FUNCTION_BLOCK EL_LinearAxis (* The logic of an equipment block: one holder at a time, outputs switched off before new ones go on, all off on release or abort, inputs reported when they change. Technical: LinearAxis: output values from its holder -> outputs (break before make); one holder at a time; all off on release or when the module aborts; inputs -> state channel when they change *)
  (* Standard: 61499-2 *)
  (* Version 0.1, 2026-09-28, Project contributors, AAU Smart Production Lab *)
  PACKAGE stoppering;
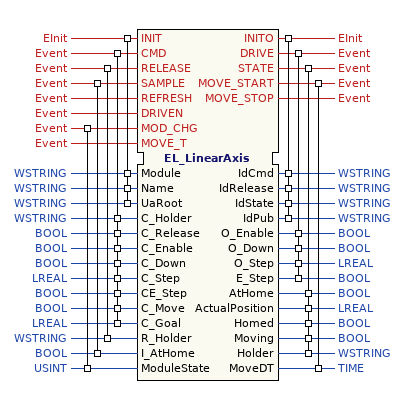
  EVENT_INPUT
    INIT : EInit WITH Module, Name, UaRoot; (* Initialise, once at start-up (the INIT chain); takes the values given with it *)
    CMD WITH C_Holder, C_Release, C_Enable, C_Down, C_Step, CE_Step, C_Move, C_Goal; (* A command arrived from a holder *)
    RELEASE WITH R_Holder; (* A release arrived on the module's release channel (R_Holder) *)
    SAMPLE WITH I_AtHome; (* The inputs were read *)
    REFRESH; (* Cycle: write the outputs again *)
    DRIVEN; (* The outputs were written *)
    MOD_CHG WITH ModuleState; (* The module's state changed (its Aborting switches all off) *)
    MOVE_T; (* The move's time is up: the axis is at the goal *)
  END_EVENT
  EVENT_OUTPUT
    INITO : EInit WITH IdCmd, IdRelease, IdState, IdPub; (* Initialised: the next block of the INIT chain goes on *)
    DRIVE WITH O_Enable, O_Down, O_Step, E_Step; (* Write the outputs *)
    STATE WITH AtHome, ActualPosition, Homed, Moving, Holder; (* Publish the state (the inputs and the holder) *)
    MOVE_START WITH MoveDT; (* Start the move's timer (MoveDT) *)
    MOVE_STOP; (* Stop the move's timer *)
  END_EVENT
  VAR_INPUT
    Module : WSTRING; (* The module's name; its local channels are named after it (loc[<Module>/...]) *)
    Name : WSTRING; (* The equipment item's name: its local channels and OPC UA folder *)
    UaRoot : WSTRING; (* The module's OPC UA folder, e.g. /Objects/Filling *)
    C_Holder : WSTRING; (* Who sends the command *)
    C_Release : BOOL; (* Give up the equipment after this command *)
    C_Enable : BOOL; (* Commanded value of Enable *)
    C_Down : BOOL; (* Commanded value of Down *)
    C_Step : LREAL; (* Commanded value of Step *)
    CE_Step : BOOL; (* Commanded: Step enabled *)
    C_Move : BOOL; (* Move to a position *)
    C_Goal : LREAL; (* The position to move to *)
    R_Holder : WSTRING; (* Who gives up the equipment *)
    I_AtHome : BOOL; (* AtHome as read or received *)
    ModuleState : USINT; (* PackML state: 1 Clearing, 2 Stopped, 3 Starting, 4 Idle, 6 Execute, 7 Stopping, 8 Aborting, 9 Aborted, 15 Resetting *)
  END_VAR
  VAR_OUTPUT
    IdCmd : WSTRING; (* Local channel of the commands *)
    IdRelease : WSTRING; (* Local channel of the releases (the module's, one for all equipment) *)
    IdState : WSTRING; (* Local channel of the state *)
    IdPub : WSTRING; (* OPC UA ID of the published inputs *)
    O_Enable : BOOL; (* The value to write to Enable *)
    O_Down : BOOL; (* The value to write to Down *)
    O_Step : LREAL; (* The value to write to Step *)
    E_Step : BOOL; (* Step enabled (FALSE writes 0) *)
    AtHome : BOOL; (* LinearAxis: AtHome, an input *)
    ActualPosition : LREAL; (* LinearAxis: ActualPosition (mm), worked out by the equipment *)
    Homed : BOOL; (* LinearAxis: Homed, worked out by the equipment *)
    Moving : BOOL; (* LinearAxis: Moving, worked out by the equipment *)
    Holder : WSTRING; (* Who holds the equipment (empty: free) *)
    MoveDT : TIME; (* How long the move takes *)
  END_VAR
  VAR
    Publish : BOOL;
    Beat : USINT;
    LastHolder : WSTRING;
    Pending : BOOL;
    OffPending : BOOL;
    L_AtHome : BOOL;
    L_Homed : BOOL;
    L_Moving : BOOL;
    N_Enable : BOOL;
    N_Down : BOOL;
    N_Step : LREAL;
    NE_Step : BOOL;
    N_Move : BOOL;
    N_Goal : LREAL;
    MoveGoal : LREAL;
    MoveFrom : LREAL;
    MoveDir : LREAL;
    MoveSince : TIME;
    MoveStart : BOOL;
    Uncounted : BOOL;
  END_VAR
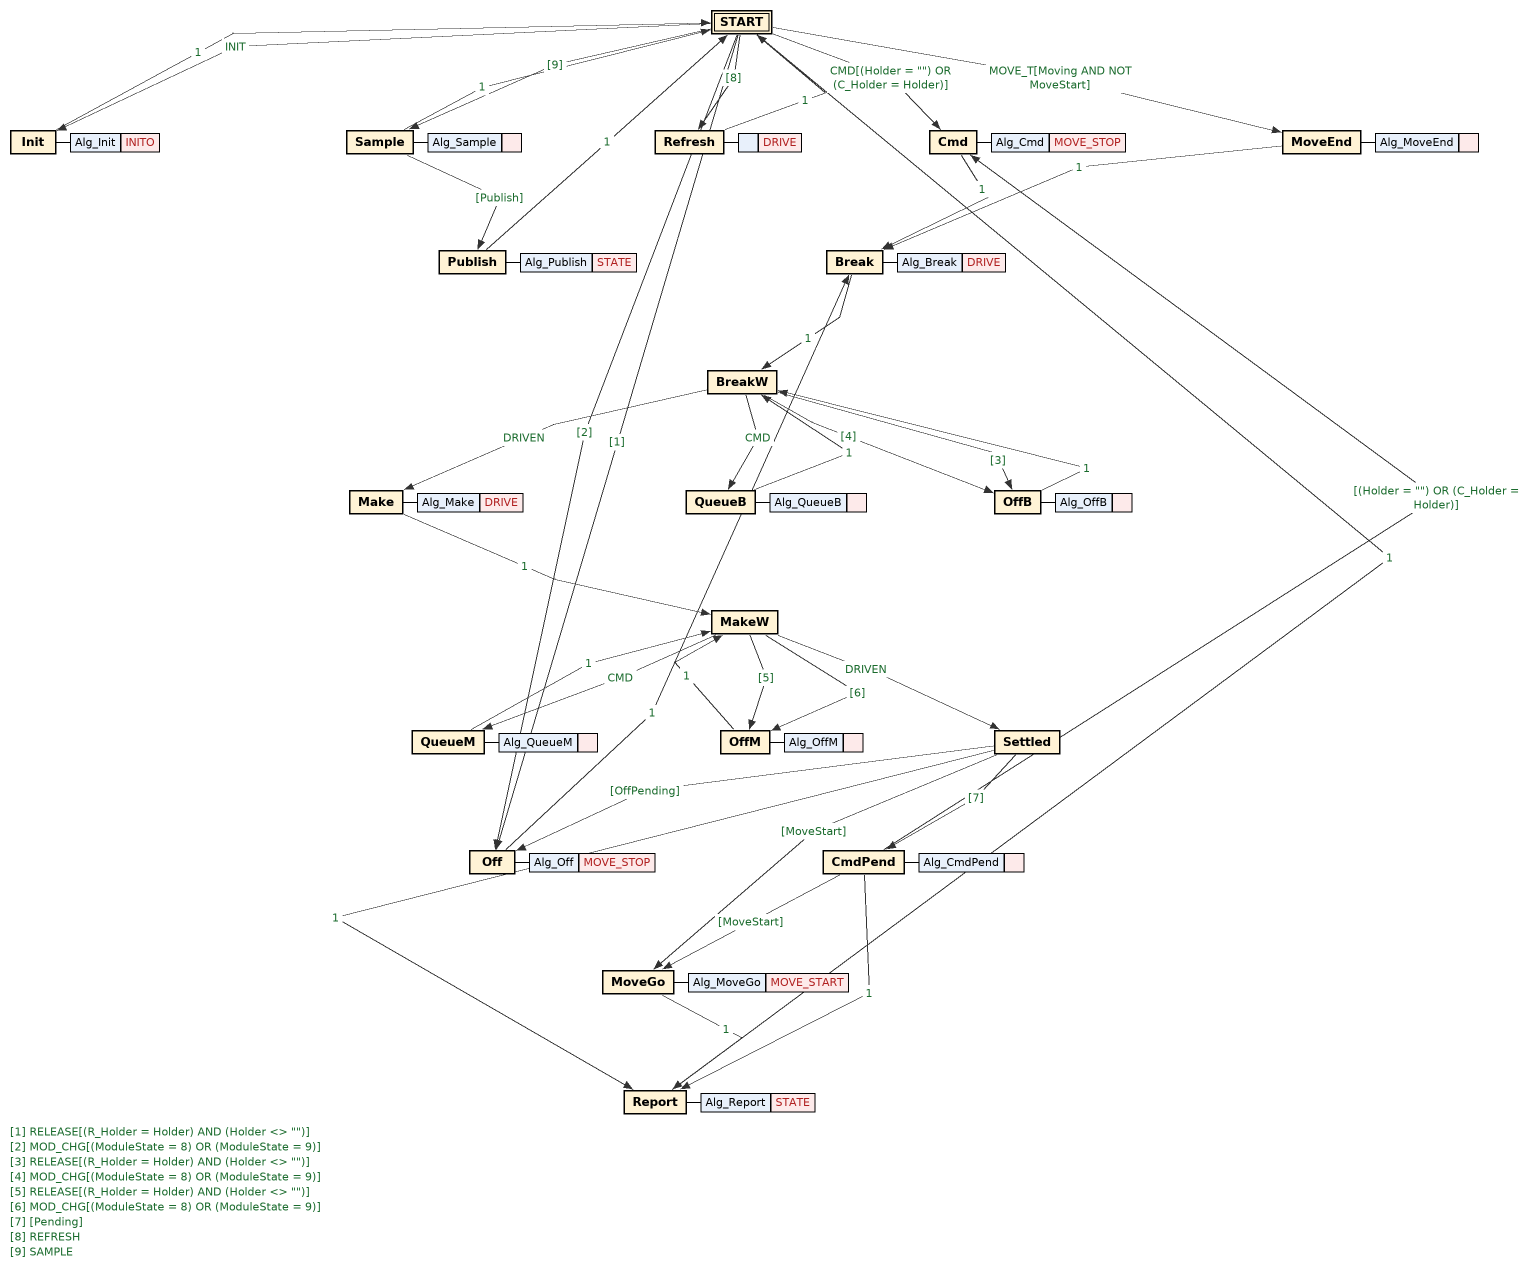
  EC_STATES
    START;
    Init : Alg_Init -> INITO;
    Sample : Alg_Sample;
    Publish : Alg_Publish -> STATE;
    Refresh : -> DRIVE;
    Cmd : Alg_Cmd -> MOVE_STOP;
    Off : Alg_Off -> MOVE_STOP;
    Break : Alg_Break -> DRIVE;
    Make : Alg_Make -> DRIVE;
    BreakW;
    MakeW;
    QueueB : Alg_QueueB;
    OffB : Alg_OffB;
    QueueM : Alg_QueueM;
    OffM : Alg_OffM;
    CmdPend : Alg_CmdPend;
    Settled;
    MoveGo : Alg_MoveGo -> MOVE_START;
    MoveEnd : Alg_MoveEnd;
    Report : Alg_Report -> STATE;
  END_STATES
  EC_TRANSITIONS
    START TO Init := INIT;
    START TO Sample := SAMPLE;
    START TO Refresh := REFRESH;
    START TO Cmd := CMD[(Holder = "") OR (C_Holder = Holder)];
    START TO Off := RELEASE[(R_Holder = Holder) AND (Holder <> "")];
    START TO Off := MOD_CHG[(ModuleState = 8) OR (ModuleState = 9)];
    START TO MoveEnd := MOVE_T[Moving AND NOT MoveStart];
    MoveEnd TO Break := 1;
    Init TO START := 1;
    Sample TO Publish := [Publish];
    Sample TO START := 1;
    Publish TO START := 1;
    Refresh TO START := 1;
    Cmd TO Break := 1;
    Off TO Break := 1;
    Break TO BreakW := 1;
    BreakW TO Make := DRIVEN;
    Make TO MakeW := 1;
    MakeW TO Settled := DRIVEN;
    BreakW TO QueueB := CMD;
    BreakW TO OffB := RELEASE[(R_Holder = Holder) AND (Holder <> "")];
    BreakW TO OffB := MOD_CHG[(ModuleState = 8) OR (ModuleState = 9)];
    QueueB TO BreakW := 1;
    OffB TO BreakW := 1;
    MakeW TO QueueM := CMD;
    MakeW TO OffM := RELEASE[(R_Holder = Holder) AND (Holder <> "")];
    MakeW TO OffM := MOD_CHG[(ModuleState = 8) OR (ModuleState = 9)];
    QueueM TO MakeW := 1;
    OffM TO MakeW := 1;
    Settled TO Off := [OffPending];
    Settled TO CmdPend := [Pending];
    CmdPend TO Cmd := [(Holder = "") OR (C_Holder = Holder)];
    CmdPend TO MoveGo := [MoveStart];
    Settled TO MoveGo := [MoveStart];
    MoveGo TO Report := 1;
    CmdPend TO Report := 1;
    Settled TO Report := 1;
    Report TO START := 1;
  END_TRANSITIONS
  ALGORITHM Alg_Init IN ST:
IdCmd := CONCAT(CONCAT(CONCAT(CONCAT("loc[", Module), "/"), Name), "/cmd]");
IdRelease := CONCAT(CONCAT("loc[", Module), "/release]");
IdState := CONCAT(CONCAT(CONCAT(CONCAT("loc[", Module), "/"), Name), "/state]");
IdPub := CONCAT(CONCAT(CONCAT(CONCAT(CONCAT(CONCAT(CONCAT(CONCAT(CONCAT(CONCAT(CONCAT(CONCAT(CONCAT(CONCAT(CONCAT(CONCAT(CONCAT("opc_ua[WRITE;", UaRoot), "/Equipment/"), Name), "/AtHome;"), UaRoot), "/Equipment/"), Name), "/ActualPosition;"), UaRoot), "/Equipment/"), Name), "/Homed;"), UaRoot), "/Equipment/"), Name), "/Moving"), "]");
  END_ALGORITHM
  ALGORITHM Alg_Sample IN ST:
AtHome := I_AtHome;
IF Moving AND NOT MoveStart THEN
  ActualPosition := MoveFrom + MoveDir * 20.0 * TIME_IN_MS_TO_LREAL(NOW_MONOTONIC() - MoveSince) / 1000.0;
  IF MoveDir * (ActualPosition - MoveGoal) > 0.0 THEN
    ActualPosition := MoveGoal;
  END_IF;
ELSIF AtHome THEN
  ActualPosition := 0.0;
  Homed := TRUE;
ELSIF Uncounted THEN
  Homed := FALSE;
END_IF;
Publish := (AtHome <> L_AtHome) OR (Homed <> L_Homed) OR (Moving <> L_Moving) OR (Holder <> LastHolder) OR (Beat >= 20) OR (Moving AND (Beat >= 4));
Beat := Beat + 1;
  END_ALGORITHM
  ALGORITHM Alg_Publish IN ST:
L_AtHome := AtHome;
L_Homed := Homed;
L_Moving := Moving;
LastHolder := Holder;
Beat := 0;
  END_ALGORITHM
  ALGORITHM Alg_Cmd IN ST:
Holder := C_Holder;
N_Enable := C_Enable;
N_Down := C_Down;
N_Step := C_Step;
NE_Step := CE_Step;
N_Move := C_Move;
N_Goal := C_Goal;
IF Moving AND NOT MoveStart THEN
  ActualPosition := MoveFrom + MoveDir * 20.0 * TIME_IN_MS_TO_LREAL(NOW_MONOTONIC() - MoveSince) / 1000.0;
  IF MoveDir * (ActualPosition - MoveGoal) > 0.0 THEN
    ActualPosition := MoveGoal;
  END_IF;
END_IF;
Moving := FALSE;
MoveStart := FALSE;
IF N_Move THEN
  IF Homed AND (ABS(N_Goal - ActualPosition) >= 0.0005) THEN
    MoveGoal := N_Goal;
    MoveFrom := ActualPosition;
    MoveDT := MUL_TIME(T#1s, ABS(N_Goal - ActualPosition) / 20.0);
    IF N_Goal > ActualPosition THEN
      MoveDir := 1.0;
      N_Enable := TRUE;
      N_Down := TRUE;
      N_Step := 50.0;
      NE_Step := TRUE;
    ELSE
      MoveDir := -1.0;
      N_Enable := TRUE;
      N_Down := FALSE;
      N_Step := 50.0;
      NE_Step := TRUE;
    END_IF;
    Moving := TRUE;
    MoveStart := TRUE;
  ELSE
    N_Enable := FALSE;
    N_Down := FALSE;
    N_Step := 0.0;
    NE_Step := FALSE;
  END_IF;
  Uncounted := FALSE;
ELSE
  Uncounted := N_Enable OR N_Down OR NE_Step;
END_IF;
IF C_Release THEN
  Holder := "";
END_IF;
  END_ALGORITHM
  ALGORITHM Alg_Off IN ST:
N_Enable := FALSE;
N_Down := FALSE;
N_Step := 0.0;
NE_Step := FALSE;
N_Move := FALSE;
N_Goal := 0.0;
IF Moving AND NOT MoveStart THEN
  ActualPosition := MoveFrom + MoveDir * 20.0 * TIME_IN_MS_TO_LREAL(NOW_MONOTONIC() - MoveSince) / 1000.0;
  IF MoveDir * (ActualPosition - MoveGoal) > 0.0 THEN
    ActualPosition := MoveGoal;
  END_IF;
END_IF;
Moving := FALSE;
MoveStart := FALSE;
Uncounted := FALSE;
Holder := "";
OffPending := FALSE;
  END_ALGORITHM
  ALGORITHM Alg_Break IN ST:
O_Enable := O_Enable AND N_Enable;
O_Down := O_Down AND N_Down;
  END_ALGORITHM
  ALGORITHM Alg_Make IN ST:
O_Enable := N_Enable;
O_Down := N_Down;
O_Step := N_Step;
E_Step := NE_Step;
  END_ALGORITHM
  ALGORITHM Alg_QueueB IN ST:
Pending := TRUE;
  END_ALGORITHM
  ALGORITHM Alg_OffB IN ST:
OffPending := TRUE;
  END_ALGORITHM
  ALGORITHM Alg_QueueM IN ST:
Pending := TRUE;
  END_ALGORITHM
  ALGORITHM Alg_OffM IN ST:
OffPending := TRUE;
  END_ALGORITHM
  ALGORITHM Alg_CmdPend IN ST:
Pending := FALSE;
  END_ALGORITHM
  ALGORITHM Alg_MoveGo IN ST:
MoveStart := FALSE;
MoveSince := NOW_MONOTONIC();
  END_ALGORITHM
  ALGORITHM Alg_MoveEnd IN ST:
ActualPosition := MoveGoal;
Moving := FALSE;
N_Enable := FALSE;
N_Down := FALSE;
N_Step := 0.0;
NE_Step := FALSE;
  END_ALGORITHM
  ALGORITHM Alg_Report IN ST:
LastHolder := Holder;
Beat := 0;
  END_ALGORITHM
END_FUNCTION_BLOCK
